Fanuc KAREL source: kt00296.KL

-- PROVISIONAL review KL for V1013-1; original PC SHA256 8247213a48fba9ef2e694ca2bc8cbc5ce380df0de8896dd5bfbc84b450aab5b2
-- Incomplete behavior may be omitted. Consult companion uncertainty JSON. Do not deploy.
PROGRAM KT00296
%NOLOCKGROUP
VAR
  I1 : INTEGER
  OUT : BOOLEAN
-- UNRESOLVED_DECL H2 type=002017
BEGIN
  -- UNRESOLVED_PC offsets 5-16; opcodes 2E,23
  -- UNRESOLVED_PC offsets 21-35; opcodes 2E,22,9D,33,B4
  -- UNRESOLVED_PC offsets 40-62; opcodes 21,22,9D,33,B3,58,23
  -- UNRESOLVED_PC offsets 67-71; opcodes 7F
END KT00296
